SUBAPPLICATION ValueOverriddenBySubAppInput
  (* Standard: 61499-1; Description: Copyright (c) 2026 Martin Erich Jobst This program and the accompanying materials are made available under the terms of the Eclipse Public License 2.0 which is available at https://www.eclipse.org/legal/epl-2.0/ SPDX-License-Identifier: EPL-2.0 *)
  (* Version 1.0, 2026-11-18, Martin Jobst *)
  PACKAGE lib::VarDeclaration;
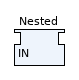
  SUBAPPLICATION Nested
    VAR_INPUT
      IN : DINT;
    END_VAR
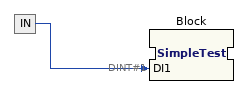
    FBS
      Block : lib::VarDeclaration::support::SimpleTest(DI1 := DINT#1);
    END_FBS
    DATA_CONNECTIONS
      IN TO Block.DI1;
    END_CONNECTIONS
  END_SUBAPPLICATION
END_SUBAPPLICATION
